SUBAPPLICATION ADI_GT_0 (* Prüft ob DINT-Adapter Wert > 0 ist (AX-Adapter Ausgang) *)
  (* Standard: 61499-2 *)
  (* Version 1.0, 2026-10-15, franz, Meisterschulen am Ostbahnhof *)
  PACKAGE MyLib::sys;
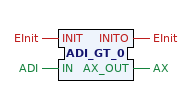
  EVENT_INPUT
    INIT : EInit; (* Initialization Request *)
  END_EVENT
  EVENT_OUTPUT
    INITO : EInit; (* Initialization Confirm *)
  END_EVENT
  SOCKETS
    IN : adapter::types::unidirectional::ADI;
  END_SOCKETS
  PLUGS
    AX_OUT : adapter::types::unidirectional::AX;
  END_PLUGS
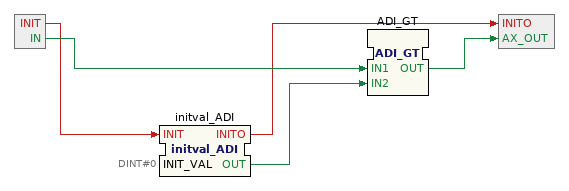
  FBS
    ADI_GT : adapter::iec61131::comparison::ADI_GT;
    initval_ADI : adapter::types::unidirectional::ADI::initval::initval_ADI(INIT_VAL := DINT#0);
  END_FBS
  EVENT_CONNECTIONS
    INIT TO initval_ADI.INIT;
    initval_ADI.INITO TO INITO;
  END_CONNECTIONS
  ADAPTER_CONNECTIONS
    IN TO ADI_GT.IN1;
    ADI_GT.OUT TO AX_OUT;
    initval_ADI.OUT TO ADI_GT.IN2;
  END_CONNECTIONS
END_SUBAPPLICATION
